FUNCTION FC 1 : VOID
BEGIN
NETWORK
      L DB1.MW 4
END_FUNCTION
